// TIA Portal V20 export
Screen "Pop-up_Opmodes24_Popup"  645x410
  ScreenItem "Background" at 0,0 size 645x410  Type=HmiRectangle
  ScreenItem "Descr_HmiPanel" at 1,350 size 56x40  Type=HmiTextBox
  ScreenItem "Linie1_LightGrey" at 10,349 size 520x0  Type=HmiLine
  ScreenItem "Linie1_DarkGrey" at 10,348 size 520x0  Type=HmiLine
  ScreenItem "Linie1_LightGrey_1" at 10,391 size 520x0  Type=HmiLine
  ScreenItem "Linie1_DarkGrey_1" at 10,390 size 520x0  Type=HmiLine
  ScreenItem "Overview_OPMode" at 1,1 size 643x25  Type=HmiTextBox
  ScreenItem "Descr_OPMode" at 1,26 size 550x40  Type=HmiTextBox
  ScreenItem "Overview_HMI-OP" at 555,350 size 90x60  Type=HmiButton
  ScreenItem "Cancel Mode" at 554,1 size 90x60  Type=HmiButton
  ScreenItem "OPMode1_small" at 15,71 size 90x60  Type=HmiButton
  ScreenItem "OPMode2_small" at 15,136 size 90x60  Type=HmiButton
  ScreenItem "OPMode3_small" at 15,201 size 90x60  Type=HmiButton
  ScreenItem "OPMode4_small" at 15,266 size 90x60  Type=HmiButton
  ScreenItem "OPMode5_small" at 122,71 size 90x60  Type=HmiButton
  ScreenItem "OPMode6_small" at 122,136 size 90x60  Type=HmiButton
  ScreenItem "OPMode7_small" at 122,201 size 90x60  Type=HmiButton
  ScreenItem "OPMode8_small" at 122,266 size 90x60  Type=HmiButton
  ScreenItem "OPMode9_small" at 226,71 size 90x60  Type=HmiButton
  ScreenItem "OPMode10_small" at 226,136 size 90x60  Type=HmiButton
  ScreenItem "OPMode11_small" at 226,201 size 90x60  Type=HmiButton
  ScreenItem "OPMode12_small" at 226,266 size 90x60  Type=HmiButton
  ScreenItem "OPMode13_small" at 331,71 size 90x60  Type=HmiButton
  ScreenItem "OPMode14_small" at 331,136 size 90x60  Type=HmiButton
  ScreenItem "OPMode15_small" at 331,201 size 90x60  Type=HmiButton
  ScreenItem "OPMode16_small" at 331,266 size 90x60  Type=HmiButton
  ScreenItem "OPMode17_small" at 435,71 size 90x60  Type=HmiButton
  ScreenItem "OPMode18_small" at 435,136 size 90x60  Type=HmiButton
  ScreenItem "OPMode19_small" at 435,201 size 90x60  Type=HmiButton
  ScreenItem "OPMode20_small" at 435,266 size 90x60  Type=HmiButton
  ScreenItem "OPMode21_smal" at 540,71 size 90x60  Type=HmiButton
  ScreenItem "OPMode22_small" at 540,136 size 90x60  Type=HmiButton
  ScreenItem "OPMode23_small" at 540,201 size 90x60  Type=HmiButton
  ScreenItem "OPMode24_small" at 540,266 size 90x60  Type=HmiButton
  ScreenItem "OPMode1_wide" at 10,71 size 100x60  Type=HmiButton
  ScreenItem "OPMode2_wide" at 10,136 size 100x60  Type=HmiButton
  ScreenItem "OPMode3_wide" at 10,201 size 100x60  Type=HmiButton
  ScreenItem "OPMode4_wide" at 10,266 size 100x60  Type=HmiButton
  ScreenItem "OPMode5_wide" at 117,71 size 100x60  Type=HmiButton
  ScreenItem "OPMode6_wide" at 117,136 size 100x60  Type=HmiButton
  ScreenItem "OPMode7_wide" at 117,201 size 100x60  Type=HmiButton
  ScreenItem "OPMode8_wide" at 117,266 size 100x60  Type=HmiButton
  ScreenItem "OPMode9_wide" at 221,71 size 100x60  Type=HmiButton
  ScreenItem "OPMode10_wide" at 221,136 size 100x60  Type=HmiButton
  ScreenItem "OPMode11_wide" at 221,201 size 100x60  Type=HmiButton
  ScreenItem "OPMode12_wide" at 221,266 size 100x60  Type=HmiButton
  ScreenItem "OPMode13_wide" at 326,71 size 100x60  Type=HmiButton
  ScreenItem "OPMode14_wide" at 326,136 size 100x60  Type=HmiButton
  ScreenItem "OPMode15_wide" at 326,201 size 100x60  Type=HmiButton
  ScreenItem "OPMode16_wide" at 326,266 size 100x60  Type=HmiButton
  ScreenItem "OPMode17_wide" at 430,71 size 100x60  Type=HmiButton
  ScreenItem "OPMode18_wide" at 430,136 size 100x60  Type=HmiButton
  ScreenItem "OPMode19_wide" at 430,201 size 100x60  Type=HmiButton
  ScreenItem "OPMode20_wide" at 430,266 size 100x60  Type=HmiButton
  ScreenItem "OPMode21_wide" at 535,71 size 100x60  Type=HmiButton
  ScreenItem "OPMode22_wide" at 535,136 size 100x60  Type=HmiButton
  ScreenItem "OPMode23_wide" at 535,201 size 100x60  Type=HmiButton
  ScreenItem "OPMode24_wide" at 535,266 size 100x60  Type=HmiButton
  ScreenItem "OPMode1_Foreground_Blocked" at 10,71 size 100x60  Type=HmiGraphicView
  ScreenItem "OPMode2_Foreground_Blocked" at 10,136 size 100x60  Type=HmiGraphicView
  ScreenItem "OPMode3_Foreground_Blocked" at 10,201 size 100x60  Type=HmiGraphicView
  ScreenItem "OPMode4_Foreground_Blocked" at 10,266 size 100x60  Type=HmiGraphicView
  ScreenItem "OPMode8_Foreground_Blocked" at 117,266 size 100x60  Type=HmiGraphicView
  ScreenItem "OPMode7_Foreground_Blocked" at 117,201 size 100x60  Type=HmiGraphicView
  ScreenItem "OPMode6_Foreground_Blocked" at 117,136 size 100x60  Type=HmiGraphicView
  ScreenItem "OPMode5_Foreground_Blocked" at 117,71 size 100x60  Type=HmiGraphicView
  ScreenItem "OPMode9_Foreground_Blocked" at 221,71 size 100x60  Type=HmiGraphicView
  ScreenItem "OPMode10_Foreground_Blocked" at 221,136 size 100x60  Type=HmiGraphicView
  ScreenItem "OPMode11_Foreground_Blocked" at 221,201 size 100x60  Type=HmiGraphicView
  ScreenItem "OPMode12_Foreground_Blocked" at 221,266 size 100x60  Type=HmiGraphicView
  ScreenItem "OPMode16_Foreground_Blocked" at 326,266 size 100x60  Type=HmiGraphicView
  ScreenItem "OPMode15_Foreground_Blocked" at 326,201 size 100x60  Type=HmiGraphicView
  ScreenItem "OPMode14_Foreground_Blocked" at 326,136 size 100x60  Type=HmiGraphicView
  ScreenItem "OPMode13_Foreground_Blocked" at 326,71 size 100x60  Type=HmiGraphicView
  ScreenItem "OPMode17_Foreground_Blocked" at 430,71 size 100x60  Type=HmiGraphicView
  ScreenItem "OPMode18_Foreground_Blocked" at 430,136 size 100x60  Type=HmiGraphicView
  ScreenItem "OPMode19_Foreground_Blocked" at 430,201 size 100x60  Type=HmiGraphicView
  ScreenItem "OPMode20_Foreground_Blocked" at 430,266 size 100x60  Type=HmiGraphicView
  ScreenItem "OPMode24_Foreground_Blocked" at 535,266 size 100x60  Type=HmiGraphicView
  ScreenItem "OPMode23_Foreground_Blocked" at 535,201 size 100x60  Type=HmiGraphicView
  ScreenItem "OPMode22_Foreground_Blocked" at 535,136 size 100x60  Type=HmiGraphicView
  ScreenItem "OPMode21_Foreground_Blocked" at 535,71 size 100x60  Type=HmiGraphicView
  ScreenItem "OPMode21_Blocked" at 616,74 size 14x14  Type=HmiGraphicView
  ScreenItem "OPMode17_Blocked" at 512,74 size 14x14  Type=HmiGraphicView
  ScreenItem "OPMode18_Blocked" at 512,140 size 14x14  Type=HmiGraphicView
  ScreenItem "OPMode19_Blocked" at 512,205 size 14x14  Type=HmiGraphicView
  ScreenItem "OPMode22_Blocked" at 616,140 size 14x14  Type=HmiGraphicView
  ScreenItem "OPMode23_Blocked" at 616,205 size 14x14  Type=HmiGraphicView
  ScreenItem "OPMode24_Blocked" at 616,270 size 14x14  Type=HmiGraphicView
  ScreenItem "OPMode20_Blocked" at 512,270 size 14x14  Type=HmiGraphicView
  ScreenItem "OPMode16_Blocked" at 406,270 size 14x14  Type=HmiGraphicView
  ScreenItem "OPMode15_Blocked" at 406,205 size 14x14  Type=HmiGraphicView
  ScreenItem "OPMode14_Blocked" at 406,140 size 14x14  Type=HmiGraphicView
  ScreenItem "OPMode13_Blocked" at 406,74 size 14x14  Type=HmiGraphicView
  ScreenItem "OPMode9_Blocked" at 304,74 size 14x14  Type=HmiGraphicView
  ScreenItem "OPMode10_Blocked" at 304,140 size 14x14  Type=HmiGraphicView
  ScreenItem "OPMode11_Blocked" at 304,205 size 14x14  Type=HmiGraphicView
  ScreenItem "OPMode12_Blocked" at 304,270 size 14x14  Type=HmiGraphicView
  ScreenItem "OPMode8_Blocked" at 200,270 size 14x14  Type=HmiGraphicView
  ScreenItem "OPMode7_Blocked" at 200,205 size 14x14  Type=HmiGraphicView
  ScreenItem "OPMode6_Blocked" at 200,140 size 14x14  Type=HmiGraphicView
  ScreenItem "OPMode5_Blocked" at 200,74 size 14x14  Type=HmiGraphicView
  ScreenItem "OPMode1_Blocked" at 93,74 size 14x14  Type=HmiGraphicView
  ScreenItem "OPMode2_Blocked" at 93,140 size 14x14  Type=HmiGraphicView
  ScreenItem "OPMode3_Blocked" at 93,205 size 14x14  Type=HmiGraphicView
  ScreenItem "OPMode4_Blocked" at 93,270 size 14x14  Type=HmiGraphicView
